(* IEC 61131-3 sources: SRCI_CLIENT_PLC/RobotLibrary/Library/Structures/AxesGroup/Parameter/Rob, 3 files *)

(* ---- AxesGroupParameterRob.st ---- *)
{attribute 'pack_mode' := '1'}
// -------------------------------------------------------------------------
//  SRCI Robot Library
// -------------------------------------------------------------------------
//
//  Object:      AxesGroupParameterRob
//  Author:      Thorsten Brach
//  Date:        2024-06-01
//
//  Description:
//
//
//  Copyright:
//    (C) 2024 Thorsten Brach. All rights reserved
//             Licensed under the MIT License.
//
//  Disclaimer:
//    This project is provided without any guarantee and can be used for
//    private and commercial purposes. Any use is at the user’s
//    own risk and responsibility.
//
// -------------------------------------------------------------------------
TYPE AxesGroupParameterRob :
STRUCT
  /// Parameter
  Parameter      : AxesGroupParameterRobParameter;
  /// Optional cyclic
  OptionalCyclic : AxesGroupParameterRobOptionalCyclic;
END_STRUCT
END_TYPE

(* ---- AxesGroupParameterRobOptionalCyclic.st ---- *)
{attribute 'pack_mode' := '1'}
// -------------------------------------------------------------------------
//  SRCI Robot Library
// -------------------------------------------------------------------------
//
//  Object:      AxesGroupParameterOptionalCyclicRobToPlc
//  Author:      Thorsten Brach
//  Date:        2024-06-01
//
//  Description:
//
//
//  Copyright:
//    (C) 2024 Thorsten Brach. All rights reserved
//             Licensed under the MIT License.
//
//  Disclaimer:
//    This project is provided without any guarantee and can be used for
//    private and commercial purposes. Any use is at the user’s
//    own risk and responsibility.
//
// -------------------------------------------------------------------------
TYPE AxesGroupParameterRobOptionalCyclic :
STRUCT
  /// Bit 00:
  /// Transmit cyclic data from PLC to RC for the usage in a subprogram on the RC called via the function “CallSubprogram”
  UseCallSubprogram       : BOOL;
  /// Bit 01:
  /// Send a short cartesian position with TCP position (X, Y,Z), rotation (RX, RY, RZ),
  /// configuration bytes (Config, TurnNumber), position of first external axis (E1) and corresponding coordinate systems (ToolNo, FrameNo)
  UseCartesianPosition    : BOOL;
  /// Bit 02:
  /// Send a short axes position with joint values (J1, J2, J3, J4, J5, J6) and position of first external axis (E1)
  UseJointPosition        : BOOL;
  /// Bit 03:
  /// Send the force with the divided forces in the individual directions (X, Y, Z, RX, RY, RZ)
  UseForce                : BOOL;
  /// Bit 04:
  /// Transmit actual axes current of individual axes (J1, J2, J3, J4, J5, J6)
  UseCurrent              : BOOL;
  /// Bit 05:
  Bit05                   : BOOL;
  /// Bit 06:
  Bit06                   : BOOL;
  /// Bit 07:
  Bit07                   : BOOL;
  /// Bit 08:
  /// Set to 1 to define two Sequences in one Telegram.
  /// If activated, 2 sequences also has to be activated in the ServerClient direction
  UseTwoSequences         : BOOL;
  /// Bit 09:
  /// Send the external axis values for an extended cartesian position (E2, E3, E4, E5, E6)
  UseCartesianPositionExt : BOOL;
  /// Bit 10:
  /// Send the external axis values for an extended joint position (E2, E3, E4, E5, E6)
  UseJointPositionExt     : BOOL;
  /// Bit 11:
  /// Transmit the current force for the external axis (E1, E2, E3, E4, E5, E6)
  UseForceExt             : BOOL;
  /// Bit 12:
  /// Transmit the actual current for the external axis (E1, E2, E3, E4, E5, E6)
  UseCurrentExt           : BOOL;
  /// Bit 13:
  Bit13                   : BOOL;
  /// Bit 14:
  Bit14                   : BOOL;
  /// Bit 15:
  Bit15                   : BOOL;
END_STRUCT
END_TYPE

(* ---- AxesGroupParameterRobParameter.st ---- *)
{attribute 'pack_mode' := '1'}
// -------------------------------------------------------------------------
//  SRCI Robot Library
// -------------------------------------------------------------------------
//
//  Object:      AxesGroupParameterRob
//  Author:      Thorsten Brach
//  Date:        2024-06-01
//
//  Description:
//
//
//  Copyright:
//    (C) 2024 Thorsten Brach. All rights reserved
//             Licensed under the MIT License.
//
//  Disclaimer:
//    This project is provided without any guarantee and can be used for
//    private and commercial purposes. Any use is at the user’s
//    own risk and responsibility.
//
// -------------------------------------------------------------------------
TYPE AxesGroupParameterRobParameter :
STRUCT
  /// User defined robot name
  RobotName                 : STRING(20);
  /// Returns a metric of how many CMDs it can receive and manage at the same time
  /// must be initialized with a value > 3, because during the interface initialization at least 3 commands are executed
  /// after ReadRobotData command the value is set to the correct ACR length wich is supported by the RC.
  LengthACR                 : UINT := 50;
  /// Highest index of available tools on the RC.
  HighestToolIndex          : USINT;
  /// Highest index of available frames on the RC.
  HighestFrameIndex         : USINT;
  /// Highest index of available loads on the RC.
  HighestLoadIndex          : USINT;
  /// Highest index of available work areas on the RC.
  HighestWorkAreaIndex      : USINT;
  /// Datas which are synchronized
  DataInSync                : DataInSync;
  /// Index of tool changed on RC
  ChangeIndexTool           : USINT;
  /// Index of frame changed on RC
  ChangeIndexFrame          : USINT;
  /// Index of load changed on RC
  ChangeIndexLoad           : USINT;
  ///Index of work area changed on RC
  ChangeIndexWorkArea       : USINT;
  /// Working hours of an RA connected to the RC
  RAWorkingHours            : UDINT;
  /// Signals that a brake test is required in the defined monitoring time (see chapter 6.5.27)
  BrakeTestRequired         : BOOL;
  /// StepMode is active and set to ExactStop (see chapter 6.1.3)
  StepModeExactStopActive   : BOOL;
  /// StepMode is active and set to Blending (see chapter 6.1.3)
  StepModeBlendingActive    : BOOL;
  /// PathAccuracyMode is active (see chapter 6.5.22)
  PathAccuracyMode          : BOOL;
  /// AvoidSingularity is active (see chapter 6.5.23)
  AvoidSingularity          : BOOL;
  /// CollisionDetection is active (see chapter 6.5.35)
  CollisionDetectionEnabled : BOOL;
  /// Cyclic dynamics status bit Accelerating is supported by RC (see chapter 5.5.3.2)
  AcceleratingSupported     : BOOL;
  /// Cyclic dynamics status bit Decelerating is supported by RC (see chapter 5.5.3.2)
  DecceleratingSupported    : BOOL;
  /// Cyclic dynamics status bit ConstantVelocity is supported by RC (see chapter 5.5.3.2)
  ConstantVelocitySupported : BOOL;
  /// Total system hours of an RA connected to the RC. Must not be modifiable by the user.
  /// •  0: Invalid
  /// • >1: Total system hours
  RCWorkingHours            : UDINT;
END_STRUCT
END_TYPE
